FUNCTION_BLOCK DrillCtrl (* Basic Function Block Type *)
  (* Standard: 61499-2 *)
  (* Version 0.0, 7/2/2026, Template *)
  PACKAGE Main;
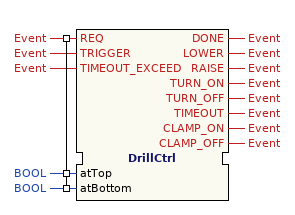
  EVENT_INPUT
    REQ WITH atTop, atBottom; (* Normal Execution Request *)
    TRIGGER;
    TIMEOUT_EXCEED;
  END_EVENT
  EVENT_OUTPUT
    DONE;
    LOWER;
    RAISE;
    TURN_ON;
    TURN_OFF;
    TIMEOUT;
    CLAMP_ON;
    CLAMP_OFF;
  END_EVENT
  VAR_INPUT
    atTop : BOOL; (* Input event qualifier *)
    atBottom : BOOL;
  END_VAR
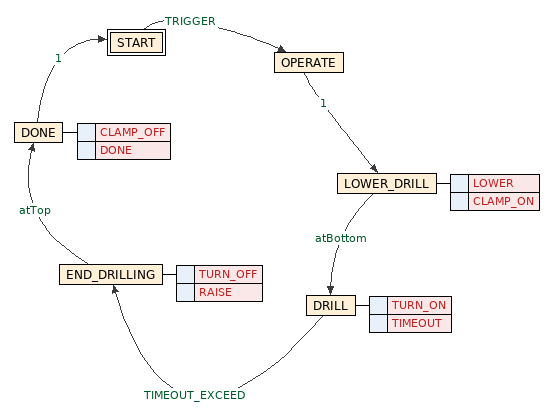
  EC_STATES
    START; (* Initial State *)
    OPERATE;
    LOWER_DRILL : -> LOWER, -> CLAMP_ON;
    DRILL : -> TURN_ON, -> TIMEOUT;
    END_DRILLING : -> TURN_OFF, -> RAISE;
    DONE : -> CLAMP_OFF, -> DONE;
  END_STATES
  EC_TRANSITIONS
    START TO OPERATE := TRIGGER;
    OPERATE TO LOWER_DRILL := 1;
    LOWER_DRILL TO DRILL := atBottom;
    DRILL TO END_DRILLING := TIMEOUT_EXCEED;
    END_DRILLING TO DONE := atTop;
    DONE TO START := 1;
  END_TRANSITIONS
  ALGORITHM INIT IN ST: (* Initialization algorithm *)
;
  END_ALGORITHM
  ALGORITHM REQ IN ST: (* Normally executed algorithm *)
;
  END_ALGORITHM
END_FUNCTION_BLOCK
